(* IEC 61131-3 sources: llm-plc-st-eval/data/processed_definitivo/qwen2.5-coder_14b/B2/zero_shot, 3 files *)

(* ---- ejec_1.st ---- *)
FUNCTION_BLOCK FB_Valvula
VAR_INPUT
    nivelAlto : BOOL; // Sensor de nivel alto
END_VAR

VAR_OUTPUT
    valvula : BOOL; // Salida para controlar la válvula
END_VAR

VAR
    timer : TON; // Timer de retardo
    estado : BOOL; // Estado de la válvula
END_VAR

// Inicialización del timer
IF timer.Q = FALSE THEN
    timer(IN := nivelAlto, PT := T#5S);
END_IF;

// Control de la válvula
IF nivelAlto THEN
    // Si el nivel está alto y el timer ha terminado, abrir la válvula
    IF timer.Q THEN
        estado := TRUE;
    END_IF;
ELSE
    // Si el nivel no está alto, cerrar la válvula inmediatamente
    estado := FALSE;
    timer(IN := FALSE); // Reiniciar el timer
END_IF;

// Asignar el estado de la válvula a la salida
valvula := estado;

(* ---- ejec_2.st ---- *)
FUNCTION_BLOCK FB_Valvula
VAR_INPUT
    nivelAlto : BOOL; // Sensor de nivel alto
END_VAR

VAR_OUTPUT
    valvula : BOOL; // Salida para controlar la válvula
END_VAR

VAR
    timer : TON; // Timer de conteo ascendente
    estado : BOOL; // Estado de la válvula
END_VAR

// Inicialización del timer
IF NOT nivelAlto THEN
    timer(IN := FALSE);
    estado := FALSE;
END_IF;

// Control de la válvula
IF nivelAlto THEN
    timer(IN := TRUE, PT := T#5S);
    IF timer.Q THEN
        estado := TRUE;
    END_IF;
ELSE
    estado := FALSE;
    timer(IN := FALSE);
END_IF;

// Asignación de la salida
valvula := estado;

(* ---- ejec_3.st ---- *)
FUNCTION_BLOCK FB_Valvula
VAR_INPUT
    nivelAlto : BOOL; // Sensor de nivel alto
END_VAR

VAR_OUTPUT
    valvula : BOOL; // Control de la válvula
END_VAR

VAR
    timer : TON; // Timer de 5 segundos
    estado : BOOL; // Estado de la válvula
END_VAR

// Inicialización del timer
IF NOT nivelAlto THEN
    timer(IN := FALSE);
    estado := FALSE;
END_IF;

// Control de la válvula
IF nivelAlto THEN
    timer(IN := TRUE);
    IF timer.Q THEN
        estado := TRUE;
    END_IF;
ELSE
    estado := FALSE;
    timer(IN := FALSE);
END_IF;

// Asignación de la salida
valvula := estado;
